(* IEC 61131-3 sources: STruCpp/tests/st-validation/variables, 6 files *)

(* ---- constants.st ---- *)
PROGRAM ConstantsTest
  VAR CONSTANT
    PI : REAL := 3.14159;
    MAX_SIZE : INT := 100;
  END_VAR
  VAR
    area : REAL;
    doubled : INT;
  END_VAR

  area := PI * 5.0 * 5.0;
  doubled := MAX_SIZE * 2;
END_PROGRAM

(* ---- initialization.st ---- *)
PROGRAM InitTest
  VAR
    init_int : INT := 42;
    init_real : REAL := 3.14;
    uninit_int : INT;
    uninit_bool : BOOL;
  END_VAR
END_PROGRAM

(* ---- test_constants.st ---- *)
TEST 'Constant REAL used in expression'
  VAR uut : ConstantsTest; END_VAR
  uut();
  ASSERT_NEAR(uut.area, 78.5397, 0.01);
END_TEST

TEST 'Constant INT used in expression'
  VAR uut : ConstantsTest; END_VAR
  uut();
  ASSERT_EQ(uut.doubled, 200);
END_TEST

(* ---- test_initialization.st ---- *)
TEST 'INT initialized to 42'
  VAR uut : InitTest; END_VAR
  ASSERT_EQ(uut.init_int, 42);
END_TEST

TEST 'REAL initialized to 3.14'
  VAR uut : InitTest; END_VAR
  ASSERT_NEAR(uut.init_real, 3.14, 0.01);
END_TEST

TEST 'Uninitialized INT defaults to 0'
  VAR uut : InitTest; END_VAR
  ASSERT_EQ(uut.uninit_int, 0);
END_TEST

TEST 'Uninitialized BOOL defaults to FALSE'
  VAR uut : InitTest; END_VAR
  ASSERT_FALSE(uut.uninit_bool);
END_TEST

(* ---- test_type_defaults.st ---- *)
TEST 'BOOL defaults to FALSE'
  VAR uut : TypeDefaultsTest; END_VAR
  ASSERT_FALSE(uut.d_bool);
END_TEST

TEST 'SINT defaults to 0'
  VAR uut : TypeDefaultsTest; END_VAR
  ASSERT_EQ(uut.d_sint, 0);
END_TEST

TEST 'INT defaults to 0'
  VAR uut : TypeDefaultsTest; END_VAR
  ASSERT_EQ(uut.d_int, 0);
END_TEST

TEST 'DINT defaults to 0'
  VAR uut : TypeDefaultsTest; END_VAR
  ASSERT_EQ(uut.d_dint, 0);
END_TEST

TEST 'USINT defaults to 0'
  VAR uut : TypeDefaultsTest; END_VAR
  ASSERT_EQ(uut.d_usint, 0);
END_TEST

TEST 'UINT defaults to 0'
  VAR uut : TypeDefaultsTest; END_VAR
  ASSERT_EQ(uut.d_uint, 0);
END_TEST

TEST 'REAL defaults to 0.0'
  VAR uut : TypeDefaultsTest; END_VAR
  ASSERT_NEAR(uut.d_real, 0.0, 0.001);
END_TEST

TEST 'LREAL defaults to 0.0'
  VAR uut : TypeDefaultsTest; END_VAR
  ASSERT_NEAR(uut.d_lreal, 0.0, 0.001);
END_TEST

(* ---- type_defaults.st ---- *)
PROGRAM TypeDefaultsTest
  VAR
    d_bool : BOOL;
    d_sint : SINT;
    d_int : INT;
    d_dint : DINT;
    d_usint : USINT;
    d_uint : UINT;
    d_real : REAL;
    d_lreal : LREAL;
  END_VAR
END_PROGRAM
